Fanuc KAREL source: kf00101.KL

-- PROVISIONAL review KL for V1013-1; original PC SHA256 4a175e20366c8bd2b8cd3ac54ef4a596dc4dde417b5deeff6f8b97c0a1a32aa5
-- Incomplete behavior may be omitted. Consult companion uncertainty JSON. Do not deploy.
PROGRAM KF00101
%NOLOCKGROUP
BEGIN
  -- UNRESOLVED_PC offsets 5-16; opcodes 2E,23
  -- UNRESOLVED_PC offsets 21-32; opcodes 2E,23
  -- UNRESOLVED_PC offsets 37-63; opcodes 27,27,9D,22,27,9D,31,7E,4A
  -- UNRESOLVED_PC offsets 68-72; opcodes 7F
END KF00101
